FUNCTION_BLOCK MotorBaseNer (* Copia do SE.App2CommonProcess.MotorBase (Schneider) com FbFail = realimentacao OU falha OU intertravamento *)
  (* Standard: 61499-2 *)
  (* Version 1.0.1, 1/30/2024, ApplicationLibDevTeam, Schneider Electric, Hidryco 04/11/2026: copia do SE.App2CommonProcess MotorBase 26.0.0.13 (export da Schneider). FbFail = AlarmStatus do feedbackFailure OU Fail OU IlckCond (FbFailCalc, FbFailComposto). Original: First Version *)
  PACKAGE SE.Nereda;
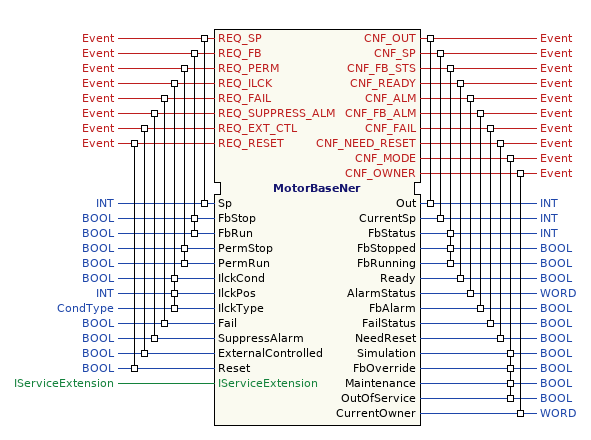
  EVENT_INPUT
    REQ_SP WITH Sp; (* Request to update setpoint *)
    REQ_FB WITH FbStop, FbRun; (* Request to update feedbacks *)
    REQ_PERM WITH PermStop, PermRun; (* Request to update permissive conditions *)
    REQ_ILCK WITH IlckCond, IlckPos, IlckType; (* Request to update interlock conditions *)
    REQ_FAIL WITH Fail; (* Request to update out of service and fail status and parameters *)
    REQ_SUPPRESS_ALM WITH SuppressAlarm; (* Request to update the alarm suppress status *)
    REQ_EXT_CTL WITH ExternalControlled; (* Request External control signal *)
    REQ_RESET WITH Reset; (* Request to reset the device *)
  END_EVENT
  EVENT_OUTPUT
    CNF_OUT WITH Out; (* Execution of confirmation output *)
    CNF_SP WITH CurrentSp; (* Execution of confirmation Current Setpoint *)
    CNF_FB_STS WITH FbRunning, FbStopped, FbStatus; (* Execution of confirmed state *)
    CNF_READY WITH Ready; (* Execution of Ready status *)
    CNF_ALM WITH AlarmStatus; (* Execution of confirmation  alarm conditions *)
    CNF_FB_ALM WITH FbAlarm; (* Execution of confirmation  Fb alarm *)
    CNF_FAIL WITH FailStatus; (* Execution of confirmation  failure *)
    CNF_NEED_RESET WITH NeedReset; (* Request for Reset *)
    CNF_MODE WITH Simulation, FbOverride, Maintenance, OutOfService; (* Excecution of new operational modes *)
    CNF_OWNER WITH CurrentOwner; (* Request for  owner *)
  END_EVENT
  VAR_INPUT
    Sp : INT; (* Setpoint of device (0 = Stop, 1 = Run,) *)
    FbStop : BOOL; (* 1 = Device stop feedback active *)
    FbRun : BOOL; (* 1 = Device run feedback active *)
    PermStop : BOOL := TRUE; (* 1 = Device stop permission active *)
    PermRun : BOOL := TRUE; (* 1 = Device run permission active *)
    IlckCond : BOOL; (* 1 = Interlock condition active *)
    IlckPos : INT; (* Interlock setpoint state (0 = Stop, 1 = Run, 3 = Interlock inactive) *)
    IlckType : CondType; (* Type of condition interlock, (0 = Normal, 1 = Process interlock/Sequence interlock) *)
    Fail : BOOL; (* 1 = Failure is active *)
    SuppressAlarm : BOOL; (* 1 = Suppress alarm in HMI *)
    ExternalControlled : BOOL; (* 1 = External control is active *)
    Reset : BOOL; (* 1 = Reset device failure *)
  END_VAR
  VAR_OUTPUT
    Out : INT; (* Calculate output of the device ( 0 = Stop command, 1 = Run command) *)
    CurrentSp : INT; (* Output value considering permissive conditions *)
    FbStatus : INT; (* Confirmed state of the device (0 = Stopped, 1 =Running, 253 = Unknown) *)
    FbStopped : BOOL; (* 1 = Stopped *)
    FbRunning : BOOL; (* 1 = Running *)
    Ready : BOOL; (* 1 = Device is ready to run *)
    AlarmStatus : WORD; (* Bit 1 = Device failure status, Bit 2 = Feedback failure status *)
    FbAlarm : BOOL; (* 1 = Feedback failure alarm is active *)
    FailStatus : BOOL; (* 1 = Fail active *)
    NeedReset : BOOL; (* 1 = Device need reset to resume the operation *)
    Simulation : BOOL; (* 1 = Simulation mode is active *)
    FbOverride : BOOL; (* 1 = Feedback overide (Sp = FbStatus) *)
    Maintenance : BOOL; (* 1 = Maintenance mode is active *)
    OutOfService : BOOL; (* 1 = Out of service mode is active *)
    CurrentOwner : WORD;
  END_VAR
  SOCKETS
    IServiceExtension : IServiceExtension(PermActive2 := TRUE, ServiceState := TRUE); (* Services extension adapter(Seq control, Local panel, Maintenance and Owner) *)
  END_SOCKETS
  (* Alarm Managment *)
  (* Control *)
  (* Data exchange with sequence *)
  (* Initialization *)
  (* Supervision Interface *)
  (* Owner & Setpoint Management *)
  FBS
    plcStart : plcStart(Delay := T#0ms, Prio := 16);
    IThis : MotorBaseNer_HMI(QI := TRUE);
    spSelection : devInSel(EnBumpless1 := FALSE, EnBumpless2 := TRUE, EnBumpless3 := FALSE, Val1 := (picosecs:=0,quality:=16#0,timestamp:=LDT#1970-01-01-05:30:00,value:=0), PermActive2 := FALSE, ResetSp := (value:=0,quality:=16#0,timestamp:=LDT#2023-01-20-10:13:38,picosecs:=0)); {SET_ATTRIBUTE(Configuration.Component.HideUnusedPorts, )}
    control : motorLogic; {SET_ATTRIBUTE(Configuration.Component.HideUnusedPorts, )}
    basicOwner : ownerControl;
    deviceFailure : stateAlarmBasic(AlarmState := TRUE); {SET_ATTRIBUTE(HMI.AlarmText, Falha do equipamento)} {SET_ATTRIBUTE(Configuration.Component.HideUnusedPorts, )}
    feedbackFailure : stateAlarmBasic(AlarmState := TRUE); {SET_ATTRIBUTE(HMI.AlarmText, Falha de realimentação: ligado/desligado não confirmado)} {SET_ATTRIBUTE(Configuration.Component.HideUnusedPorts, )}
    progSpSelection : SELECT_24363B89CFDE21263; {SET_ATTRIBUTE(Configuration.GenericFBType.InterfaceParams, Runtime.Standard#CNT:=2;SELECT:BOOL;IN${CNT$}:INT)}
    resetConditions : DS_SELECTX_1579ED5B8ACDFC94C; {SET_ATTRIBUTE(Configuration.GenericFBType.InterfaceParams, Runtime.Standard#CNTX:=3;CNTY:=1;DI${CNTX,_,CNTY$}:BOOL)}
    FbFailCalc : FbFailComposto;
  END_FBS
  EVENT_CONNECTIONS
    spSelection.CNF TO control.REQ_SP;
    control.CNF_OUT TO IServiceExtension.CNF_STATUS;
    control.CNF_FB_STS TO IServiceExtension.CNF_STATUS;
    spSelection.CNF TO IServiceExtension.CNF_STATUS;
    control.CNF_FB_ALM TO CNF_FB_ALM;
    control.CNF_READY TO IServiceExtension.CNF_READY;
    control.CNF_MODE TO IServiceExtension.CNF_OPMODE;
    REQ_SUPPRESS_ALM TO IServiceExtension.CNF_SUPPRESS_ALM;
    REQ_SUPPRESS_ALM TO deviceFailure.REQ_SUPRESS;
    control.CNF_FB_STS TO CNF_FB_STS;
    control.CNF_OUT TO CNF_OUT;
    control.CNF_MODE TO CNF_MODE;
    REQ_FB TO control.REQ_FB;
    REQ_ILCK TO control.REQ_ILCK;
    REQ_FAIL TO control.REQ_FAIL;
    deviceFailure.INITO TO feedbackFailure.INIT;
    REQ_PERM TO spSelection.REQ_SEL;
    IServiceExtension.REQ_OWNER TO basicOwner.REQ_STDOWNER;
    basicOwner.CNF_OWNER TO spSelection.REQ_SEL;
    feedbackFailure.INITO TO plcStart.ACK_FIRST;
    control.CNF_NEED_RESET TO CNF_NEED_RESET;
    control.CNF_READY TO CNF_READY;
    spSelection.CNF TO CNF_SP;
    REQ_EXT_CTL TO control.REQ_EXT_CTL;
    control.CNF_FAIL TO deviceFailure.REQ;
    control.CNF_FAIL TO CNF_FAIL;
    plcStart.FIRST_INIT TO IThis.34A017503AC1070A;
    IThis.377462E9CE5193B5 TO IThis.F2953B6BB9388F21;
    control.CNF_FB_STS TO IThis.EC791CA6E67D66B3;
    control.CNF_OUT TO IThis.EC791CA6E67D66B3;
    control.CNF_NEED_RESET TO IThis.EC791CA6E67D66B3;
    spSelection.CNF TO IThis.EC791CA6E67D66B3;
    control.CNF_TRANS_FB TO IThis.EC791CA6E67D66B3;
    REQ_SUPPRESS_ALM TO IThis.EC791CA6E67D66B3;
    deviceFailure.CNF_ALM TO IThis.EC791CA6E67D66B3;
    feedbackFailure.CNF_ALM TO FbFailCalc.594458DF2A5BB47C;
    IThis.377462E9CE5193B5 TO deviceFailure.INIT;
    IThis.95BEA68906019444 TO control.REQ_PARA;
    IThis.C6CA4032A5F6989A TO spSelection.REQ_SP2;
    IThis.4711DA9A2DFC024 TO basicOwner.REQ_FORCE;
    IThis.4711DA9A2DFC024 TO control.REQ_PARA;
    IThis.4711DA9A2DFC024 TO spSelection.REQ_SEL;
    control.CNF_FAIL TO IThis.EC791CA6E67D66B3;
    control.CNF_ILCK TO IThis.EC791CA6E67D66B3;
    REQ_PERM TO IThis.EC791CA6E67D66B3;
    plcStart.FIRST_INIT TO IServiceExtension.CNF_SERVICE;
    control.CNF_FB_ALM TO feedbackFailure.REQ;
    IThis.95BEA68906019444 TO feedbackFailure.REQ_PARA;
    IThis.95BEA68906019444 TO deviceFailure.REQ_PARA;
    control.CNF_ALM TO CNF_ALM;
    control.CNF_ILCK TO spSelection.REQ_SEL;
    control.CNF_FAIL TO spSelection.RESET_SP;
    REQ_SUPPRESS_ALM TO feedbackFailure.REQ_SUPRESS;
    basicOwner.CNF_OWNER TO IThis.EC791CA6E67D66B3;
    IThis.B42FC414051FE233 TO basicOwner.REQ_BASICOWNER;
    IThis.377462E9CE5193B5 TO basicOwner.REQ_BASICOWNER;
    REQ_PERM TO IServiceExtension.CNF_READY;
    REQ_SP TO progSpSelection.REQ;
    IServiceExtension.REQ_CMD TO progSpSelection.REQ;
    progSpSelection.CNF TO spSelection.REQ_SP3;
    control.CNF_ALM TO IServiceExtension.CNF_READY;
    control.CNF_ILCK TO IServiceExtension.CNF_READY;
    REQ_EXT_CTL TO IThis.EC791CA6E67D66B3;
    basicOwner.CNF_OWNER TO CNF_OWNER;
    REQ_RESET TO resetConditions.REQ3;
    IServiceExtension.REQ_RESET TO resetConditions.REQ2;
    IThis.1A2B085F4B246BF1 TO resetConditions.REQ1;
    resetConditions.IND TO control.REQ_RESET;
    control.CNF_NEED_RESET TO IServiceExtension.CNF_READY;
    IThis.95BEA68906019444 TO IServiceExtension.CNF_CFG;
    FbFailCalc.16943D7D3AD410BC TO IThis.EC791CA6E67D66B3;
    REQ_FAIL TO FbFailCalc.594458DF2A5BB47C;
    REQ_ILCK TO FbFailCalc.594458DF2A5BB47C;
  END_CONNECTIONS
  DATA_CONNECTIONS
    spSelection.PermVal TO control.Sp;
    control.FbStatus TO IServiceExtension.Status;
    spSelection.PermVal TO IServiceExtension.CurrentSp;
    control.Out TO IServiceExtension.CurrentOp;
    control.NeedReset TO IServiceExtension.NeedReset;
    control.FbAlarm TO FbAlarm;
    control.Mode TO IServiceExtension.OpMode;
    control.Ready TO IServiceExtension.Ready;
    SuppressAlarm TO IServiceExtension.SuppressAlarm;
    SuppressAlarm TO deviceFailure.Suppress;
    SuppressAlarm TO feedbackFailure.Suppress;
    control.FbAlarm TO feedbackFailure.Input;
    control.FailStatus TO FailStatus;
    IlckPos TO control.IlckPos;
    IlckCond TO control.IlckCond;
    IlckType TO control.IlckType;
    FbStop TO control.FbStop;
    FbRun TO control.FbRun;
    Fail TO control.Fail;
    PermStop TO spSelection.PermPassive;
    PermRun TO spSelection.PermActive1;
    control.FbStopped TO FbStopped;
    control.FbRunning TO FbRunning;
    control.Out TO Out;
    control.FbStatus TO FbStatus;
    basicOwner.ProgramOwner TO spSelection.Sel3;
    basicOwner.OperatorOwner TO spSelection.Sel2;
    IlckPos TO spSelection.IlckSp;
    control.Interlocked TO spSelection.Ilck;
    IServiceExtension.StdOwner TO basicOwner.StdOwner;
    control.NeedReset TO NeedReset;
    control.Ready TO Ready;
    ExternalControlled TO control.ExternalControlled;
    control.FailStatus TO deviceFailure.Input;
    control.FbStatus TO IThis.E35507CB164A688E;
    control.TransFbStatus TO IThis.937CA40F4D16204B;
    control.Out TO IThis.D2C35BC47DF71FCC;
    spSelection.PermVal TO IThis.C6876D790F3A950E;
    control.NeedReset TO IThis.9CD6749867E91606;
    feedbackFailure.AlarmStatus TO FbFailCalc.3F9FEFE8A07BE74F;
    deviceFailure.AlarmStatus TO IThis.E4BB2C7DF94BE70A;
    control.Interlocked TO IThis.22A0744EA4DC0124;
    IThis.922C4AB423622B98 TO basicOwner.BasicOwner;
    IThis.861B8773AF2757FC TO control.MonTime;
    IThis.5568E3E91B9AAED8 TO control.TripTime;
    IThis.22AB1FF8E4CF2F97 TO control.FailResetReq;
    IThis.869E02415F6A841 TO spSelection.Val2;
    IThis.CF1EA84FDDBF53A1 TO control.Simulation;
    IThis.CF1EA84FDDBF53A1 TO Simulation;
    IThis.AD38F01F8F0043E7 TO control.FbOverride;
    IThis.AD38F01F8F0043E7 TO FbOverride;
    IThis.C8DEEF765E4F14C0 TO basicOwner.ForceOperator;
    IThis.C8DEEF765E4F14C0 TO Maintenance;
    IThis.6EDFC17C06F3153 TO control.OutOfService;
    IThis.6EDFC17C06F3153 TO spSelection.Sel1;
    IThis.152A2BD44E46F288 TO deviceFailure.ScanTime;
    IThis.152A2BD44E46F288 TO feedbackFailure.ScanTime;
    IThis.3CCC10520A21214A TO deviceFailure.AckType;
    IThis.3CCC10520A21214A TO feedbackFailure.AckType;
    IThis.89CD17990DC40B0E TO spSelection.EnTrackSp;
    IThis.B2B61A4BABE50F70 TO spSelection.EnResetSp;
    PermStop TO IThis.AB1D2B96094C90BD;
    basicOwner.StdOwnerConnected TO IThis.621B2EAA60B4DCF6;
    IThis.C8DEEF765E4F14C0 TO control.Maintenance;
    control.AlarmStatus TO AlarmStatus;
    IThis.6EDFC17C06F3153 TO OutOfService;
    spSelection.PermVal TO CurrentSp;
    control.FailStatus TO spSelection.Fail;
    basicOwner.Owner TO IThis.9CB24E1B5B149DBC;
    PermRun TO IThis.18DA785EF50AD374;
    PermStop TO IServiceExtension.PermPassive;
    PermRun TO IServiceExtension.PermActive1;
    control.AlarmStatus TO IServiceExtension.Alarm;
    control.Interlocked TO IServiceExtension.Interlocked;
    IThis.3DA6D0F9276D43A4 TO control.ConfResetReq;
    basicOwner.StdOwnerConnected TO progSpSelection.SELECT;
    Sp TO progSpSelection.IN1;
    IServiceExtension.Sp TO progSpSelection.IN2;
    progSpSelection.OUT TO spSelection.Val3;
    ExternalControlled TO IThis.130A3A1CA20AF67A;
    basicOwner.Owner TO CurrentOwner;
    Reset TO resetConditions.DI3_1;
    IServiceExtension.Reset TO resetConditions.DI2_1;
    IThis.4D34C1A4533BA5DF TO resetConditions.DI1_1;
    resetConditions.OUT1 TO control.Reset;
    IThis.89CD17990DC40B0E TO IServiceExtension.EnTrackSp;
    IThis.B2B61A4BABE50F70 TO IServiceExtension.EnResetSp;
    control.Failure TO IThis.D28866DFD0C1393B;
    FbFailCalc.CA70046049C9A2EC TO IThis.7F794E74835A9A2;
    IlckCond TO FbFailCalc.C72C731F987D59D4;
    Fail TO FbFailCalc.12594D80635DBCE8;
  END_CONNECTIONS
END_FUNCTION_BLOCK
